// TIA Portal V21 export
FUNCTION "FC_AnaTempRead" : Int   // FC10, SCL
TITLE = Analyzer: Temp read before written
{ S7_Optimized_Access := 'TRUE' }
// Rule C26c: Sum is read before it is written
// stored: SetENOAutomatically false
   VAR_INPUT
      Value : Int;   // Value to add
   END_VAR
   VAR_TEMP
      Sum : Int;   // Temporary sum
   END_VAR
BEGIN

       #Sum := #Sum + #Value;
       #FC_AnaTempRead := #Sum;
END_FUNCTION
